(* CODESYS project jsontools.library
   DefaultNamespace: KOSTAL.AF2024.Core.JsonTools
   DocFormat: reStructuredText
   Description: Base functionalities to handle a json File
   Author: Frank Dümpelmann
   Title: KOSTAL.AF2024.Core.JsonTools
   Version: 1.0.0.0
   Company: KOSTAL GmbH & Co.KG
   Placeholder: KOSTAL.AF2024.Core.JsonTools

Project tree, tasks and I/O mapping:
  libraries: KOSTAL.AF2024.Core.Process, 1.0.0.0 (KOSTAL GmbH & Co.KG); KOSTAL.AF2024.Core.Settings, 1.0.0.0 (KOSTAL GmbH & Co.KG); KOSTAL.AF2024.Core.StringTools, 1.0.0.0 (KOSTAL GmbH & Co.KG); KOSTAL.AF2024.Core.System, 1.0.0.0 (KOSTAL GmbH & Co.KG); Tc2_Standard, 3.3.3.0 (Beckhoff Automation GmbH); Tc2_System, 3.6.2.0 (Beckhoff Automation GmbH); Tc2_Utilities, 3.5.2.0 (Beckhoff Automation GmbH); Tc3_IotBase, 3.3.2.0 (Beckhoff Automation GmbH); Tc3_JsonXml, 3.4.3.0 (Beckhoff Automation GmbH)
  0_Core/
    function block _FB_Core [ST]: _DocumentIsEmpty, _FBmain, _GetArrayElementByIndex, _GetArraySize, _GetDocument, _GetDocumentLenght, _NewDocument, FB_exit, FBmain
  1_Base/
    0_Protected/
      function block _FB_Base_PE [ST]: _ReadExtStorage, _ReadFileStorage, _FB_Main_EXT, _Step_ClearContent, _Step_CreateContent, _Step_Idle_EXT, _Step_ParseContent, _Step_ReadFile, _Step_ValidateFile, _Step_WriteFileAs, _Step_WriteFileVerification, _Step_Clear, _Step_failed, _Step_Finish, _Step_FinishFail, _Step_Idle, _Step_ValidateParameter, _WriteExtAsStorage, _wFV_a0_ChainFail, _wFV_a0_Finish, _wFV_a10_Origin, _wFV_a10_Read, _WriteFileAsStorage, _extStorageDefine, _FBmain, _PE_Ex_ReadExt, _PE_Ex_ReadFile, _PE_Ex_SaveFileAs, _PE_Ex_SaveToExtAs, _PE_Clear, _PE_FBmain
    1_Public/
      0_Fundamental/
        function block _FB_Base [ST]: Clear, FBmain, LinkExtStorage, extFileName, extFilePath, fullQualifiedFile, State, TimeOut
      1_DataSourceAccess/
        function block _FB_Base_RO [ST]: Ex_ReadExt, Ex_ReadFile
        function block _FB_Base_RW [ST]: Ex_SaveFileAs, Ex_SaveToExtAs, Retries
  DUT/
    data type E_THIS_CALLED
  PARSING/
    function block _FB_Parsing [ST]: PARSE_ARRAY, PARSE_BOOL, PARSE_BYTE, PARSE_DINT, PARSE_JSON, PARSE_LREAL, PARSE_MEMBER, PARSE_REAL, PARSE_STRING, PARSE_TIME, PARSE_UDINT, PARSE_ULINT
    function block _FB_Parsing_PE [ST]: _PARSE_ARRAY, _PARSE_BOOL, _PARSE_BYTE, _PARSE_DINT, _PARSE_JSON, _PARSE_LREAL, _PARSE_MEMBER, _PARSE_REAL, _PARSE_STRING, _PARSE_TIME, _PARSE_UDINT, _PARSE_ULINT
  Project Information/
    function F_GetCompany [ST]
    function F_GetTitle [ST]
    function F_GetVersion [ST]
  Storage/
    interface I_JsonStorage: Ex_Read, Ex_Write, LinkJsonParser, State
  Version/
    global variables Global_Version
*)

// DUT/E_THIS_CALLED
{attribute 'qualified_only'}
{attribute 'strict'}
TYPE E_THIS_CALLED :
(
	IDL := 0,
	FILE_READ,
	FILE_WRITE,
	WEB_READ,
	WEB_WRITE,
	CLEAR
);
END_TYPE

// Version/Global_Version
{attribute 'TcGenerated'}
{attribute 'no-analysis'}
{attribute 'linkalways'}
// This function has been automatically generated from the project information.
VAR_GLOBAL CONSTANT
	{attribute 'const_non_replaced'}
	stLibVersion_KOSTAL_AF2024_Core_JsonTools : ST_LibVersion := (iMajor := 1, iMinor := 0, iBuild := 0, iRevision := 0, nFlags := 0, sVersion := '1.0.0.0');
END_VAR

// 0_Core/_FB_Core
(*
	Use the FB_Core class if you want to use your own json data source.
	e.g. a STRING(4096) on a communication.
*)
FUNCTION_BLOCK ABSTRACT _FB_Core EXTENDS _FB_Parsing_PE

VAR
	
	_jDoc		: Tc3_IotBase.SJsonValue;	

	_concat	: Kostal_AF2024_Core_StringTools.FB_CONCAT;
	
END_VAR

VAR CONSTANT
	_EMPTY_DOC_LENGHT	: UDINT:= 5;
END_VAR

METHOD PROTECTED _DocumentIsEmpty : BOOL

_DocumentIsEmpty:= _parser.GetDocumentLength() <= _EMPTY_DOC_LENGHT;
END_METHOD

METHOD PROTECTED _FBmain : BOOL
;
END_METHOD

METHOD PROTECTED _GetArrayElementByIndex : Tc3_IotBase.SJsonValue
VAR_INPUT
	jContainer	: Tc3_IotBase.SJsonValue;
	Index				: UDINT;
	state				: REFERENCE TO KOSTAL_AF2024_Core_Settings.T_MaxString;		
END_VAR

VAR
	_state					: KOSTAL_AF2024_Core_Settings.T_MaxString;	
END_VAR
IF jContainer = 0 THEN _state:= "GetArraySize - jContainer Parameter is empty";	

ELSIF Index >= _parser.GetArraySize(jContainer) THEN	_state:= "GetArraySize - Index is out of range";

ELSE	_GetArrayElementByIndex:= _parser.GetArrayValueByIdx(jContainer, Index);

END_IF

IF __ISVALIDREF(state) THEN state:= _state;	END_IF
END_METHOD

METHOD PROTECTED _GetArraySize : UDINT;
VAR_INPUT
	jContainer	: Tc3_IotBase.SJsonValue;
	state				: REFERENCE TO KOSTAL_AF2024_Core_Settings.T_MaxString;		
END_VAR

VAR
	_state	: KOSTAL_AF2024_Core_Settings.T_MaxString;	
END_VAR
IF jContainer = 0 THEN _state:= "GetArraySize - jContainer Parameter is empty";	

ELSE	_GetArraySize:= _parser.GetArraySize(jContainer);
	
END_IF

IF __ISVALIDREF(state) THEN state:= _state;	END_IF
END_METHOD

(*
getDocument
===========

|return a Pointer >Tc3_IotBase.SJsonValue< to jason document
*)

METHOD PROTECTED _GetDocument : Tc3_IotBase.SJsonValue;
_GetDocument:= _jDoc;
END_METHOD

METHOD PROTECTED _GetDocumentLenght : UDINT;
VAR_INPUT
END_VAR
_GetDocumentLenght:= _parser.GetDocumentLength();
END_METHOD

(*
use in your _Step_CreateContent to start with an empty json File
*)
METHOD PROTECTED _NewDocument : BOOL

_parser.NewDocument();

_jDoc:= _parser.GetDocumentRoot();

_GetDocumentLenght();

_NewDocument:= _jDoc <> 0;
END_METHOD

METHOD FB_exit : BOOL
VAR_INPUT
	bInCopyCode : BOOL; // if TRUE, the exit method is called for exiting an instance that is copied afterwards (online change).
END_VAR

_NewDocument();
END_METHOD

METHOD PUBLIC FBmain
VAR_INPUT
END_VAR
;
END_METHOD

END_FUNCTION_BLOCK

// PARSING/_FB_Parsing_PE
(*
	Contains protected methods to parse various data types.
*)
FUNCTION_BLOCK ABSTRACT _FB_Parsing_PE

VAR
	_parser	: Tc3_JsonXml.FB_JsonDomParser;
END_VAR

(*
Returns the Json Array Element of jContainer
*)
METHOD PROTECTED _PARSE_ARRAY : Tc3_IotBase.SJsonValue;

VAR_INPUT
	jContainer	: Tc3_IotBase.SJsonValue;
	Member			: KOSTAL_AF2024_Core_Settings.T_MaxString_UTF8;	
	mustExist		: BOOL;
	state				: REFERENCE TO KOSTAL_AF2024_Core_Settings.T_MaxString_UTF8;		
END_VAR

VAR
	_J						:	Tc3_IotBase.SJsonValue;
	_state	: KOSTAL_AF2024_Core_Settings.T_MaxString_UTF8;	
END_VAR
_PARSE_ARRAY:= 0;
_state:= '';

IF jContainer = 0 																		THEN	_state:= Tc2_Standard.CONCAT(Member,  ';PARSE_ARRAY - jContainer Parameter is empty');	

ELSIF NOT _parser.HasMember(jContainer, Member)	THEN	_state:= Tc2_Standard.CONCAT(Member,  ';PARSE_ARRAY - no member');

ELSE

	_J:= _parser.FindMember(jContainer,	Member);

	IF _J = 0 										THEN 	_state:= Tc2_Standard.CONCAT(Member,  ';PARSE_ARRAY - no member');	
	ELSIF _parser.IsNull(_J)	THEN 	_state:= Tc2_Standard.CONCAT(Member,  ';PARSE_ARRAY - is NULL');	
	ELSE																_PARSE_ARRAY:= _J;
	END_IF

END_IF

IF __ISVALIDREF(state) THEN state:= _state;	END_IF
END_METHOD

(*
Returns a bool Value of jContainer
*)
METHOD PROTECTED _PARSE_BOOL : BOOL

VAR_INPUT
	jContainer	: Tc3_IotBase.SJsonValue;
	Member			: KOSTAL_AF2024_Core_Settings.T_MaxString_UTF8;	
	mustExist		: BOOL;
	state				: REFERENCE TO KOSTAL_AF2024_Core_Settings.T_MaxString_UTF8;		
END_VAR

VAR
	_J			:	Tc3_IotBase.SJsonValue;
	_state	: KOSTAL_AF2024_Core_Settings.T_MaxString_UTF8;	
END_VAR
_PARSE_BOOL:= FALSE; 
_state:= '';

IF jContainer = 0 THEN _state:= Tc2_Standard.CONCAT(Member,  ';PARSE_BOOL - jContainer Parameter is empty');

ELSIF NOT _parser.HasMember(jContainer, Member) THEN
	
	IF mustExist THEN	_state:= Tc2_Standard.CONCAT(Member,  ';PARSE_BOOL - no member');	END_IF

ELSE

	_J:= _parser.FindMember(jContainer,	Member);

	IF _J = 0 											THEN	IF mustExist	THEN	_state:= Tc2_Standard.CONCAT(Member,  ';PARSE_BOOL - no member');	END_IF
	ELSIF _parser.IsNull(_J)		THEN	IF mustExist	THEN	_state:= Tc2_Standard.CONCAT(Member,  ';PARSE_BOOL - is NULL');	END_IF
	ELSIF _parser.IsBool(_J)		THEN	_PARSE_BOOL:= _parser.GetBool(v:= _J);	
	ELSIF _parser.IsNumber(_J)	THEN	_PARSE_BOOL:=  UDINT_TO_BOOL(_parser.GetUint(_J));
	ELSIF _parser.IsString(_J)	THEN	_PARSE_BOOL:=  STRING_TO_BOOL(_parser.GetString(_J));
	ELSE																	IF mustExist 	THEN	_state:= Tc2_Standard.CONCAT(Member,  ';PARSE_BOOL - not BOOL');	END_IF
	END_IF

END_IF
	
IF __ISVALIDREF(state) THEN state:= _state;	END_IF
END_METHOD

(*
Returns a byte Value of jContainer
*)
METHOD PROTECTED _PARSE_BYTE : BYTE

VAR_INPUT
	jContainer	: Tc3_IotBase.SJsonValue;
	Member			: KOSTAL_AF2024_Core_Settings.T_MaxString_UTF8;	
	mustExist		: BOOL;
	state				: REFERENCE TO KOSTAL_AF2024_Core_Settings.T_MaxString_UTF8;		
END_VAR

VAR
	_J						:	Tc3_IotBase.SJsonValue;
	_state				: KOSTAL_AF2024_Core_Settings.T_MaxString_UTF8;	
END_VAR
_PARSE_BYTE:= 0; 
_state:= '';

IF jContainer = 0 THEN _state:= Tc2_Standard.CONCAT(Member,  ';PARSE_BYTE - jContainer Parameter is empty');

ELSIF NOT _parser.HasMember(jContainer, Member) THEN
	
	IF mustExist THEN	_state:= Tc2_Standard.CONCAT(Member,  ';PARSE_BYTE - no member');	END_IF

ELSE

	_J:= _parser.FindMember(jContainer,	Member);

	IF _J = 0 											THEN	IF mustExist	THEN	_state:= Tc2_Standard.CONCAT(Member,  ';PARSE_BYTE - no member');	END_IF
	ELSIF _parser.IsNull(_J)		THEN	IF mustExist	THEN	_state:= Tc2_Standard.CONCAT(Member,  ';PARSE_BYTE - is NULL');	END_IF
	ELSIF _parser.IsBool(_J)		THEN	_PARSE_BYTE:= 	BOOL_TO_BYTE(_parser.GetBool(v:= _J));	
	ELSIF _parser.IsNumber(_J)	THEN	_PARSE_BYTE:=  UDINT_TO_BYTE(_parser.GetUint(_J));
	ELSIF _parser.IsString(_J)	THEN	_PARSE_BYTE:=  STRING_TO_BYTE(_parser.GetString(_J));
	ELSE																	IF mustExist 	THEN	_state:= Tc2_Standard.CONCAT(Member,  ';PARSE_BYTE - not BYTE');	END_IF
	END_IF

END_IF
	
IF __ISVALIDREF(state) THEN state:= _state;	END_IF
END_METHOD

(*
Returns a DINT Value of jContainer
*)
METHOD PROTECTED _PARSE_DINT : DINT

VAR_INPUT
	jContainer	: Tc3_IotBase.SJsonValue;
	Member			: KOSTAL_AF2024_Core_Settings.T_MaxString_UTF8;	
	mustExist		: BOOL;
	state				: REFERENCE TO KOSTAL_AF2024_Core_Settings.T_MaxString_UTF8;		
END_VAR

VAR
	_J						:	Tc3_IotBase.SJsonValue;
	_state				: KOSTAL_AF2024_Core_Settings.T_MaxString_UTF8;	
END_VAR
_PARSE_DINT:= 0; 
_state:= '';

IF jContainer = 0 THEN _state:= Tc2_Standard.CONCAT(Member,  ';PARSE_DINT - jContainer Parameter is empty');

ELSIF NOT _parser.HasMember(jContainer, Member) THEN
	
	IF mustExist THEN	_state:= Tc2_Standard.CONCAT(Member,  ';PARSE_DINT - no member');	END_IF

ELSE

	_J:= _parser.FindMember(jContainer,	Member);

	IF _J = 0 											THEN	IF mustExist	THEN	_state:= Tc2_Standard.CONCAT(Member,  ';PARSE_DINT - no member');	END_IF
	ELSIF _parser.IsNull(_J)		THEN	IF mustExist	THEN	_state:= Tc2_Standard.CONCAT(Member,  ';PARSE_DINT - is NULL');	END_IF
	ELSIF _parser.IsBool(_J)		THEN	_PARSE_DINT:= 	BOOL_TO_DINT(_parser.GetBool(v:= _J));	
	ELSIF _parser.IsNumber(_J)	THEN	_PARSE_DINT:=  UDINT_TO_DINT(_parser.GetUint(_J));
	ELSIF _parser.IsString(_J)	THEN	_PARSE_DINT:=  STRING_TO_DINT(_parser.GetString(_J));
	ELSE																	IF mustExist 	THEN	_state:= Tc2_Standard.CONCAT(Member,  ';PARSE_DINT - not DINT');	END_IF
	END_IF

END_IF
	
IF __ISVALIDREF(state) THEN state:= _state;	END_IF
END_METHOD

(*
Returns the Json Element of jContainer
*)
METHOD PROTECTED _PARSE_JSON : Tc3_IotBase.SJsonValue;

VAR_INPUT
	jContainer	: Tc3_IotBase.SJsonValue;
	Member			: KOSTAL_AF2024_Core_Settings.T_MaxString_UTF8;	
	mustExist		: BOOL;
	state				: REFERENCE TO KOSTAL_AF2024_Core_Settings.T_MaxString_UTF8;		
END_VAR

VAR
	_J	:	Tc3_IotBase.SJsonValue;
	_state	: KOSTAL_AF2024_Core_Settings.T_MaxString_UTF8;	
END_VAR
_PARSE_JSON:= 0;
_state:= '';

IF jContainer = 0 																		THEN	_state:= Tc2_Standard.CONCAT(Member,  ';PARSE_JSON - jContainer Parameter is empty');	

ELSIF NOT _parser.HasMember(jContainer, Member)	THEN	_state:= Tc2_Standard.CONCAT(Member,  ';PARSE_JSON - no member');

ELSE

	_J:= _parser.FindMember(jContainer,	Member);

	IF _J = 0 									THEN 	_state:= Tc2_Standard.CONCAT(Member,  ';PARSE_JSON - no member');	
	ELSIF _parser.IsNull(_J)		THEN 	_state:= Tc2_Standard.CONCAT(Member,  ';PARSE_JSON - is NULL');	
	ELSE															_PARSE_JSON:= _J;
	END_IF

END_IF

IF __ISVALIDREF(state) THEN state:= _state;	END_IF
END_METHOD

(*
Returns a ULINT Value of jContainer
*)
METHOD PROTECTED _PARSE_LREAL : LREAL

VAR_INPUT
	jContainer	: Tc3_IotBase.SJsonValue;
	Member			: KOSTAL_AF2024_Core_Settings.T_MaxString_UTF8;	
	mustExist		: BOOL;
	state				: REFERENCE TO KOSTAL_AF2024_Core_Settings.T_MaxString_UTF8;		
END_VAR

VAR
	_J						:	Tc3_IotBase.SJsonValue;
	_state				: KOSTAL_AF2024_Core_Settings.T_MaxString_UTF8;	
END_VAR

_PARSE_LREAL:= LREAL#0; 

_state:= '';

IF jContainer = 0 THEN _state:= Tc2_Standard.CONCAT(Member,  ';PARSE_LREAL - jContainer Parameter is empty');

ELSIF NOT _parser.HasMember(jContainer, Member) THEN
	
	IF mustExist THEN	_state:= Tc2_Standard.CONCAT(Member,  ';PARSE_LREAL - no member');	END_IF

ELSE

	_J:= _parser.FindMember(jContainer,	Member);

	IF _J = 0 											THEN	IF mustExist	THEN	_state:= Tc2_Standard.CONCAT(Member,  ';PARSE_LREAL - no member');	END_IF
	ELSIF _parser.IsNull(_J)		THEN	IF mustExist	THEN	_state:= Tc2_Standard.CONCAT(Member,  ';PARSE_LREAL - is NULL');	END_IF
	ELSIF _parser.IsBool(_J)		THEN	_PARSE_LREAL:= 	BOOL_TO_LREAL(_parser.GetBool(v:= _J));	
	ELSIF _parser.IsNumber(_J)	THEN	_PARSE_LREAL:= 	_parser.GetDouble(_J);
	ELSIF _parser.IsString(_J)	THEN	_PARSE_LREAL:=	STRING_TO_LREAL(_parser.GetString(_J));
	ELSE																	IF mustExist 	THEN	_state:= Tc2_Standard.CONCAT(Member,  ';PARSE_LREAL - not BYTE');	END_IF
	END_IF

END_IF
	
IF __ISVALIDREF(state) THEN state:= _state;	END_IF
END_METHOD

(*
Returns the Json Element of jContainer
*)
METHOD PROTECTED _PARSE_MEMBER : Tc3_IotBase.SJsonValue;

VAR_INPUT
	jContainer	: Tc3_IotBase.SJsonValue;
	Member			: KOSTAL_AF2024_Core_Settings.T_MaxString_UTF8;	
	mustExist		: BOOL;
	state				: REFERENCE TO KOSTAL_AF2024_Core_Settings.T_MaxString_UTF8;		
END_VAR

VAR
	_J	:	Tc3_IotBase.SJsonValue;
	_state	: KOSTAL_AF2024_Core_Settings.T_MaxString_UTF8;	
END_VAR
_PARSE_MEMBER:= 0;
_state:= '';

IF jContainer = 0 																		THEN	_state:= Tc2_Standard.CONCAT(Member,  ';PARSE_JSON - jContainer Parameter is empty');	

ELSIF NOT _parser.HasMember(jContainer, Member)	THEN	_state:= Tc2_Standard.CONCAT(Member,  ';PARSE_JSON - no member');

ELSE

	_J:= _parser.FindMember(jContainer,	Member);

	IF _J = 0																	THEN 	_state:= Tc2_Standard.CONCAT(Member,  ';PARSE_JSON - no member');
	ELSIF		mustExist AND _parser.IsNull(_J)	THEN 	_state:= Tc2_Standard.CONCAT(Member,  ';PARSE_MEMBER - is NULL');	
	ELSE																						_PARSE_MEMBER:= _J;
	END_IF

END_IF

IF __ISVALIDREF(state) THEN state:= _state;	END_IF
END_METHOD

(*
Returns a ULINT Value of jContainer
*)
METHOD PROTECTED _PARSE_REAL : REAL

VAR_INPUT
	jContainer	: Tc3_IotBase.SJsonValue;
	Member			: KOSTAL_AF2024_Core_Settings.T_MaxString_UTF8;	
	mustExist		: BOOL;
	state				: REFERENCE TO KOSTAL_AF2024_Core_Settings.T_MaxString_UTF8;		
END_VAR

VAR
	_J						:	Tc3_IotBase.SJsonValue;
	_state				: KOSTAL_AF2024_Core_Settings.T_MaxString_UTF8;	
END_VAR

_PARSE_REAL:= REAL#0; 

_state:= '';

IF jContainer = 0 THEN _state:= Tc2_Standard.CONCAT(Member,  ';PARSE_REAL - jContainer Parameter is empty');

ELSIF NOT _parser.HasMember(jContainer, Member) THEN
	
	IF mustExist THEN	_state:= Tc2_Standard.CONCAT(Member,  ';PARSE_REAL - no member');	END_IF

ELSE

	_J:= _parser.FindMember(jContainer,	Member);

	IF _J = 0 											THEN	IF mustExist	THEN	_state:= Tc2_Standard.CONCAT(Member,  ';PARSE_REAL - no member');	END_IF
	ELSIF _parser.IsNull(_J)		THEN	IF mustExist	THEN	_state:= Tc2_Standard.CONCAT(Member,  ';PARSE_REAL - is NULL');	END_IF
	ELSIF _parser.IsBool(_J)		THEN	_PARSE_REAL:= 	BOOL_TO_REAL(_parser.GetBool(v:= _J));	
	ELSIF _parser.IsNumber(_J)	THEN	_PARSE_REAL:= 	LREAL_TO_REAL(_parser.GetDouble(_J));
	ELSIF _parser.IsString(_J)	THEN	_PARSE_REAL:=	STRING_TO_REAL(_parser.GetString(_J));
	ELSE																	IF mustExist 	THEN	_state:= Tc2_Standard.CONCAT(Member,  ';PARSE_REAL - not BYTE');	END_IF
	END_IF

END_IF
	
IF __ISVALIDREF(state) THEN state:= _state;	END_IF
END_METHOD

(*
Returns a STRING Value of jContainer
*)
METHOD PROTECTED _PARSE_STRING : KOSTAL_AF2024_Core_Settings.T_MaxString_UTF8

VAR_INPUT
	jContainer	: Tc3_IotBase.SJsonValue;
	Member			: KOSTAL_AF2024_Core_Settings.T_MaxString_UTF8;	
	mustExist		: BOOL;
	state				: REFERENCE TO KOSTAL_AF2024_Core_Settings.T_MaxString_UTF8;		
END_VAR

VAR
	_J						:	Tc3_IotBase.SJsonValue;
	_state				: KOSTAL_AF2024_Core_Settings.T_MaxString_UTF8;	
END_VAR
_PARSE_STRING:= ''; 
_state:= '';

IF jContainer = 0 THEN _state:= Tc2_Standard.CONCAT(Member,  ';PARSE_STRING - jContainer Parameter is empty');

ELSIF NOT _parser.HasMember(jContainer, Member) THEN
	
	IF mustExist THEN	_state:= Tc2_Standard.CONCAT(Member,  ';PARSE_STRING - no member');	END_IF

ELSE

	_J:= _parser.FindMember(jContainer,	Member);

	IF _J = 0 									THEN	IF mustExist		THEN	_state:= Tc2_Standard.CONCAT(Member,  ';PARSE_STRING - no member');	END_IF
	ELSIF _parser.IsNull(_J)		THEN	IF mustExist		THEN	_state:= Tc2_Standard.CONCAT(Member,  ';PARSE_STRING - is NULL');	END_IF
	ELSIF _parser.IsBool(_J)		THEN	_PARSE_STRING:= 	BOOL_TO_STRING(_parser.GetBool(v:= _J));	
	ELSIF _parser.IsNumber(_J)	THEN	_PARSE_STRING:=  UDINT_TO_STRING(_parser.GetUint(_J));
	ELSIF _parser.IsString(_J)	THEN	_PARSE_STRING:=  _parser.GetString(_J);
	ELSE				IF mustExist 		THEN	_state:= Tc2_Standard.CONCAT(Member,  ';PARSE_STRING - not STRING');	END_IF
	END_IF

END_IF
	
IF __ISVALIDREF(state) THEN state:= _state;	END_IF
END_METHOD

(*
Returns a TIME Value of jContainer
*)
METHOD PROTECTED _PARSE_TIME : TIME

VAR_INPUT
	jContainer	: Tc3_IotBase.SJsonValue;
	Member			: KOSTAL_AF2024_Core_Settings.T_MaxString_UTF8;	
	mustExist		: BOOL;
	state				: REFERENCE TO KOSTAL_AF2024_Core_Settings.T_MaxString_UTF8;		
END_VAR

VAR
	_J						:	Tc3_IotBase.SJsonValue;
	_num					: ULINT;
	_state				: KOSTAL_AF2024_Core_Settings.T_MaxString_UTF8;	
END_VAR
_PARSE_TIME:= T#0MS; 
_state:= '';

IF jContainer = 0 THEN _state:= Tc2_Standard.CONCAT(Member,  ';PARSE_TIME - jContainer Parameter is empty');

ELSIF NOT _parser.HasMember(jContainer, Member) THEN
	
	IF mustExist THEN	_state:= Tc2_Standard.CONCAT(Member,  ';PARSE_TIME - no member');	END_IF

ELSE

	_J:= _parser.FindMember(jContainer,	Member);

	IF _J = 0 									THEN	IF mustExist	THEN	_state:= Tc2_Standard.CONCAT(Member,  ';PARSE_TIME - no member');	END_IF
	ELSIF _parser.IsNull(_J)		THEN	IF mustExist	THEN	_state:= Tc2_Standard.CONCAT(Member,  ';PARSE_TIME - is NULL');	END_IF
	ELSIF _parser.IsNumber(_J)	THEN	_PARSE_TIME:=  ULINT_TO_TIME(_parser.GetUint(_J));
	ELSIF _parser.IsString(_J)	THEN	_PARSE_TIME:=  STRING_TO_TIME(_parser.GetString(_J));
	ELSE					IF mustExist 	THEN	_state:= Tc2_Standard.CONCAT(Member,  ';PARSE_TIME - not BYTE');	END_IF
	END_IF

END_IF
	
IF __ISVALIDREF(state) THEN state:= _state;	END_IF
END_METHOD

(*
Returns a UDINT Value of jContainer
*)
METHOD PROTECTED _PARSE_UDINT : UDINT

VAR_INPUT
	jContainer	: Tc3_IotBase.SJsonValue;
	Member			: KOSTAL_AF2024_Core_Settings.T_MaxString_UTF8;	
	mustExist		: BOOL;
	state				: REFERENCE TO KOSTAL_AF2024_Core_Settings.T_MaxString_UTF8;		
END_VAR

VAR
	_J						:	Tc3_IotBase.SJsonValue;
	_state				: KOSTAL_AF2024_Core_Settings.T_MaxString_UTF8;	
END_VAR
_PARSE_UDINT:= 0; 
_state:= '';

IF jContainer = 0 THEN _state:= Tc2_Standard.CONCAT(Member,  ';PARSE_UDINT - jContainer Parameter is empty');

ELSIF NOT _parser.HasMember(jContainer, Member) THEN
	
	IF mustExist THEN	_state:= Tc2_Standard.CONCAT(Member,  ';PARSE_UDINT - no member');	END_IF

ELSE

	_J:= _parser.FindMember(jContainer,	Member);

	IF _J = 0 									THEN	IF mustExist	THEN	_state:= Tc2_Standard.CONCAT(Member,  ';PARSE_UDINT - no member');	END_IF
	ELSIF _parser.IsNull(_J)		THEN	IF mustExist	THEN	_state:= Tc2_Standard.CONCAT(Member,  ';PARSE_UDINT - is NULL');	END_IF
	ELSIF _parser.IsBool(_J)		THEN	_PARSE_UDINT:= BOOL_TO_UDINT(_parser.GetBool(v:= _J));	
	ELSIF _parser.IsNumber(_J)	THEN	_PARSE_UDINT:= _parser.GetUint(_J);
	ELSIF _parser.IsString(_J)	THEN	_PARSE_UDINT:=  STRING_TO_UDINT(_parser.GetString(_J));
	ELSE					IF mustExist 	THEN	_state:= Tc2_Standard.CONCAT(Member,  ';PARSE_UDINT - not BYTE');	END_IF
	END_IF

END_IF
	
IF __ISVALIDREF(state) THEN state:= _state;	END_IF
END_METHOD

(*
Returns a ULINT Value of jContainer
*)
METHOD PROTECTED _PARSE_ULINT : ULINT

VAR_INPUT
	jContainer	: Tc3_IotBase.SJsonValue;
	Member			: KOSTAL_AF2024_Core_Settings.T_MaxString_UTF8;	
	mustExist		: BOOL;
	state				: REFERENCE TO KOSTAL_AF2024_Core_Settings.T_MaxString_UTF8;		
END_VAR

VAR
	_J						:	Tc3_IotBase.SJsonValue;
	_state				: KOSTAL_AF2024_Core_Settings.T_MaxString_UTF8;	
END_VAR
_PARSE_ULINT:= 0; 
_state:= '';

IF jContainer = 0 THEN _state:= Tc2_Standard.CONCAT(Member,  ';PARSE_ULINT - jContainer Parameter is empty');

ELSIF NOT _parser.HasMember(jContainer, Member) THEN
	
	IF mustExist THEN	_state:= Tc2_Standard.CONCAT(Member,  ';PARSE_ULINT - no member');	END_IF

ELSE

	_J:= _parser.FindMember(jContainer,	Member);

	IF _J = 0										THEN	IF mustExist	THEN	_state:= Tc2_Standard.CONCAT(Member,  ';PARSE_ULINT - no member');	END_IF
	ELSIF _parser.IsNull(_J)		THEN	IF mustExist	THEN	_state:= Tc2_Standard.CONCAT(Member,  ';PARSE_ULINT - is NULL');	END_IF
	ELSIF _parser.IsBool(_J)		THEN	_PARSE_ULINT:= BOOL_TO_ULINT(_parser.GetBool(v:= _J));	
	ELSIF _parser.IsNumber(_J)	THEN	_PARSE_ULINT:= _parser.GetUint64(_J);
	ELSIF _parser.IsString(_J)	THEN	_PARSE_ULINT:=  STRING_TO_ULINT(_parser.GetString(_J));
	ELSE					IF mustExist 	THEN	_state:= Tc2_Standard.CONCAT(Member,  ';PARSE_ULINT - not BYTE');	END_IF
	END_IF

END_IF
	
IF __ISVALIDREF(state) THEN state:= _state;	END_IF
END_METHOD

END_FUNCTION_BLOCK

// 1_Base/0_Protected/_FB_Base_PE
(*
	All needed methods and parameters are available as protected _..._PE templates
	make in inherating class available in puclic methods and parameters
*)
FUNCTION_BLOCK ABSTRACT _FB_Base_PE EXTENDS _FB_Core

VAR
	
	_Step				: KOSTAL_AF2024_Core_process.FB_processStep_Flow;

	_State	: KOSTAL_AF2024_Core_Process.T_plcState;

	_THIS_CALLED			: E_THIS_CALLED;
	_THIS_IN_PROCESS	: E_THIS_CALLED;

	_fullQualifiedFile	: KOSTAL_AF2024_Core_Settings.T_MaxString_UTF8;

	_ExecuteLoad	: BOOL;
	_LoadSuccess	: BOOL;

	_ExecuteSave	: BOOL;
	_SaveSuccess	: BOOL;

	
	_TimeOutTimer	: Tc2_Standard.TON;
	_TimeOut			: TIME:= T#5S;
	
	_iExtStorage	: I_JsonStorage;
	_extFileName	: KOSTAL_AF2024_Core_Settings.T_MaxString_UTF8;
	_extFilePath	: KOSTAL_AF2024_Core_Settings.T_MaxString_UTF8;
	
	{region 'write file verification'}
		_wFV_Step						: KOSTAL_AF2024_Core_process.FB_processStep_Flow;
		_wFV_Retries				: UINT:= 3;
		_wFV_RetriesCounter	: UINT;
		_wFV_FFE						: Tc2_Utilities.FB_EnumFindFileEntry;
		_wFV_ParserFileSize	: ULINT;
		_wFV_FileSize				: ULINT;
	{endregion}
	
	_ADDRESS_writeFailAs: INT;

END_VAR

VAR CONSTANT
	_ADDRESS_IDLE					: INT:= 0;
	_ADDRESS_SAVE_FILE_AS	: INT:= 100;
	_ADDRESS_CLEAR				: INT:= 200;
	_ADDRESS_FINISH_FAIL	: INT:= 300;
END_VAR

METHOD PROTECTED _ReadExtStorage
VAR_INPUT
END_VAR
IF _Step.toggle THEN	

	_TimeOutTimer(IN:= FALSE);	

	IF _iExtStorage = 0 THEN
		
		_State.clear();
		_State.finish:= TRUE;
		_State.fail:= TRUE;
		_State.description:= "web storage is not linked";
		
		_Step.set(_ADDRESS_FINISH_FAIL);

		RETURN;
	
	ELSIF NOT _iExtStorage.State.ready	THEN

		_State.clear();
		_State.finish:= TRUE;
		_State.fail:= TRUE;
		_State.description:= "web storage is not ready";
		
		_Step.set(_ADDRESS_FINISH_FAIL);

		RETURN;

	END_IF
	
END_IF


_TimeOutTimer(IN:= TRUE, PT:= _TimeOut);

IF _TimeOutTimer.Q THEN

	_State.clear();
	_State.finish:= TRUE;
	_State.fail:= TRUE;
	_State.description:= "File not able to read";

	_Step.set(_ADDRESS_FINISH_FAIL);

ELSIF NOT _iExtStorage.Ex_Read(_extFileName, _extFilePath) THEN	

	_State.clear();
	_State.busy:= TRUE;
	_State.description:= Tc2_Standard.WCONCAT("wait for web call accept;", _iExtStorage.State.description);

ELSIF NOT _iExtStorage.State.finish THEN	

	_State.clear();
	_State.busy:= TRUE;
	_State.description:= Tc2_Standard.WCONCAT("wait for web response;", _iExtStorage.State.description);

ELSIF NOT _iExtStorage.State.pass THEN	

	_State.clear();
	_State.finish:= TRUE;
	_State.fail:= TRUE;
	_State.description:= Tc2_Standard.WCONCAT("web call failed;", _iExtStorage.State.description);

	_Step.set(_ADDRESS_FINISH_FAIL);

ELSE	

	_jDoc:= _parser.GetDocumentRoot();
	_Step.INC();
			
END_IF
END_METHOD

METHOD PROTECTED _ReadFileStorage
VAR_INPUT
END_VAR


IF _Step.toggle THEN	_ExecuteLoad:= TRUE; _TimeOutTimer(IN:= FALSE);	END_IF

_TimeOutTimer(IN:= _ExecuteLoad, PT:= _TimeOut);

IF _ExecuteLoad THEN
	_LoadSuccess:= _parser.LoadDocumentFromFile(_fullQualifiedFile, _ExecuteLoad);
END_IF

IF _TimeOutTimer.Q THEN

	_State.clear();
	_State.finish:= TRUE;
	_State.fail:= TRUE;
	_State.description:= "File not able to read";

ELSIF _ExecuteLoad THEN	

	_State.description:= "Wait for LoadDocument Response";

ELSIF NOT _LoadSuccess THEN	

	_State.clear();
	_State.finish:= TRUE;
	_State.fail:= TRUE;
	_State.description:= "LoadDocument failed";
	
ELSE	

	_jDoc:= _parser.GetDocumentRoot();
	_Step.INC();
			
END_IF
END_METHOD

(*
	Overwrite to add your FBmain extension
*)
METHOD PROTECTED _FB_Main_EXT : BOOL
VAR_INPUT
END_VAR
END_METHOD

(*
	Overwrite to clear your data content before parse content
*)
METHOD PROTECTED _Step_ClearContent

_Step.INC();
END_METHOD

(*
	Overwrite to create your data content
*)
METHOD PROTECTED _Step_CreateContent

_Step.INC();
END_METHOD

(*
	Overwrite to add your Idle content here
*)
METHOD PROTECTED _Step_Idle_EXT : BOOL
VAR_INPUT
END_VAR

_Step_Idle_EXT:= FALSE;
END_METHOD

(*
	Overwrite to parse your data content
*)
METHOD PROTECTED _Step_ParseContent

_Step.INC();
END_METHOD

METHOD PROTECTED _Step_ReadFile
VAR_INPUT
END_VAR

IF 		_THIS_IN_PROCESS = E_THIS_CALLED.FILE_READ 	THEN	_ReadFileStorage();
ELSIF	_THIS_IN_PROCESS = E_THIS_CALLED.WEB_READ 	THEN	_ReadExtStorage();
ELSE

	_State.clear();
	_State.description:= Tc2_Standard.WCONCAT("no valid process in _Step_ReadFile; IN_PROCESS: ", INT_TO_WSTRING(_THIS_IN_PROCESS));
	_State.finish:= TRUE;
	_State.fail:= TRUE;
	_step.set(_ADDRESS_FINISH_FAIL);

END_IF
END_METHOD

METHOD PROTECTED _Step_ValidateFile
VAR_INPUT
END_VAR

_State.clear();
_State.finish:= TRUE;

IF _DocumentIsEmpty() THEN	

	_State.clear();
	_State.finish:= TRUE;
	_State.fail:= TRUE;
	_State.description:= "File not found or empty";

ELSE

	_Step.INC();

END_IF
END_METHOD

METHOD PROTECTED _Step_WriteFileAs
VAR_INPUT
END_VAR

_ADDRESS_writeFailAs:= _Step.actual;

IF 		_THIS_IN_PROCESS = E_THIS_CALLED.FILE_WRITE THEN	_WriteFileAsStorage();
ELSIF	_THIS_IN_PROCESS = E_THIS_CALLED.WEB_WRITE 	THEN	_WriteExtAsStorage();
ELSE

	_State.clear();
	_State.description:= Tc2_Standard.WCONCAT("no valid process in _Step_WriteFileAs; IN_PROCESS: ", INT_TO_WSTRING(_THIS_IN_PROCESS));
	_State.finish:= TRUE;
	_State.fail:= TRUE;
	_step.set(_ADDRESS_FINISH_FAIL);

END_IF
END_METHOD

METHOD PROTECTED _Step_WriteFileVerification

IF _THIS_IN_PROCESS <> E_THIS_CALLED.FILE_WRITE THEN	_Step.INC();
ELSE

	IF _Step.toggle	THEN	_wFV_Step.init();	END_IF
	
	_wFV_Step.Header();
	
	IF _wFV_Step.isActive(0)	THEN	_wFV_a10_Origin();	END_IF
	IF _wFV_Step.isActive(1)	THEN	_wFV_a10_Read();		END_IF
	IF _wFV_Step.isActive(2)	THEN	_wFV_a0_Finish();		END_IF
	
	IF _wFV_Step.NotFound()	THEN _wFV_a0_ChainFail();		END_IF

END_IF
END_METHOD

METHOD PROTECTED _Step_Clear
VAR_INPUT
END_VAR

_NewDocument();	

_Step.INC();
END_METHOD

METHOD PROTECTED _Step_failed
VAR_INPUT
END_VAR

_State.clear();
_State.finish:= TRUE;
_State.fail:= TRUE;

_concat.clear();
_concat.addContent("STEP Number ");
_concat.addContent(INT_TO_WSTRING(_Step.actual));
_concat.addContent(" does not exist - PLease call Support");

_State.description:= _concat.getResult();

_concat.clear();
END_METHOD

METHOD PROTECTED _Step_Finish : BOOL
VAR_INPUT
END_VAR

_State.clear();
_State.finish:= TRUE;
_State.pass:= TRUE;

_Step_Finish:= TRUE;
END_METHOD

METHOD PROTECTED _Step_FinishFail

VAR_INST
	_description	: KOSTAL_AF2024_Core_Settings.T_MaxString;
END_VAR

IF _Step.toggle THEN _description:= _State.description;	END_IF

_state.clear(); 
_state.finish := true;
_state.fail:= TRUE;

_state.description:= _description;
END_METHOD

METHOD PROTECTED _Step_Idle
VAR_INPUT
END_VAR

VAR
	_EmptyFile: KOSTAL_AF2024_Core_Settings.T_MaxString_UTF8;
END_VAR

IF _Step.toggle THEN
	
	_EmptyFile:= '';
	
	_ExecuteLoad:= FALSE;
	_LoadSuccess:= _parser.LoadDocumentFromFile(_EmptyFile, _ExecuteLoad);
	_LoadSuccess:= FALSE;

	_ExecuteSave:= FALSE;
	_SaveSuccess:= _parser.SaveDocumentToFile(_EmptyFile, _ExecuteSave);
	_SaveSuccess:= FALSE;
	
	_wFV_RetriesCounter:= UINT#0;

END_IF

IF _Step_Idle_EXT() THEN	; //Handle extended content

ELSIF _THIS_CALLED = E_THIS_CALLED.FILE_READ THEN

	_THIS_IN_PROCESS:= _THIS_CALLED;

	_NewDocument();
	_State.clear();
	_State.busy:= TRUE;
	_step.INC();


ELSIF _THIS_CALLED = E_THIS_CALLED.WEB_READ THEN

	_THIS_IN_PROCESS:= _THIS_CALLED;
	
	_NewDocument();
	_State.clear();
	_State.busy:= TRUE;
	_step.INC();



ELSIF _THIS_CALLED = E_THIS_CALLED.FILE_WRITE THEN

	_THIS_IN_PROCESS:= _THIS_CALLED;

	_State.clear();
	_State.busy:= TRUE;
	_step.set(_ADDRESS_SAVE_FILE_AS);


ELSIF _THIS_CALLED = E_THIS_CALLED.WEB_WRITE THEN

	_THIS_IN_PROCESS:= _THIS_CALLED;

	_State.clear();
	_State.busy:= TRUE;
	_step.set(_ADDRESS_SAVE_FILE_AS);



ELSIF _THIS_CALLED = E_THIS_CALLED.CLEAR THEN

	_THIS_IN_PROCESS:= _THIS_CALLED;

	_State.clear();
	_State.busy:= TRUE;
	_step.set(_ADDRESS_CLEAR);

ELSE

	_THIS_IN_PROCESS:= E_THIS_CALLED.IDL;	

	_State.clear();
	_State.ready:= TRUE;


END_IF
END_METHOD

METHOD PROTECTED _Step_ValidateParameter
VAR_INPUT
END_VAR

IF (_THIS_IN_PROCESS = E_THIS_CALLED.FILE_READ)
OR (_THIS_IN_PROCESS = E_THIS_CALLED.FILE_WRITE) 	
THEN

	IF _fullQualifiedFile = '' THEN	

		_State.clear();
		_State.finish:= TRUE;
		_State.fail:= TRUE;
		_State.description:= "fullQualifiedFile is empty";

	ELSE

		_Step.INC();
		
	END_IF

ELSIF (_THIS_IN_PROCESS = E_THIS_CALLED.WEB_READ)
OR 		(_THIS_IN_PROCESS = E_THIS_CALLED.WEB_WRITE) 	
THEN

	IF _extFileName = '' THEN	

		_State.clear();
		_State.finish:= TRUE;
		_State.fail:= TRUE;
		_State.description:= "webFileName is empty";

	ELSIF _extFilePath = '' THEN	

		_State.clear();
		_State.finish:= TRUE;
		_State.fail:= TRUE;
		_State.description:= "webFilePath is empty";

	ELSE

		_Step.INC();
		
	END_IF

ELSE
	
	_Step.INC();

END_IF
END_METHOD

METHOD PROTECTED _WriteExtAsStorage
VAR_INPUT
END_VAR
IF _Step.toggle THEN	

	_TimeOutTimer(IN:= FALSE);	

	IF _iExtStorage = 0 THEN
		
		_State.clear();
		_State.finish:= TRUE;
		_State.fail:= TRUE;
		_State.description:= "web storage is not linked";
		
		_Step.set(_ADDRESS_FINISH_FAIL);

		RETURN;
	
	ELSIF NOT _iExtStorage.State.ready	THEN

		_State.clear();
		_State.finish:= TRUE;
		_State.fail:= TRUE;
		_State.description:= "web storage is not ready";
		
		_Step.set(_ADDRESS_FINISH_FAIL);

		RETURN;

	END_IF
	
END_IF


_TimeOutTimer(IN:= TRUE, PT:= _TimeOut);

IF _TimeOutTimer.Q THEN

	_State.clear();
	_State.finish:= TRUE;
	_State.fail:= TRUE;
	_State.description:= "File not able to write";

	_Step.set(_ADDRESS_FINISH_FAIL);

ELSIF NOT _iExtStorage.Ex_Write(_extFileName, _extFilePath) THEN	

	_State.clear();
	_State.busy:= TRUE;
	_State.description:= Tc2_Standard.WCONCAT("wait for web call accept;", _iExtStorage.State.description);

ELSIF NOT _iExtStorage.State.finish THEN	

	_State.clear();
	_State.busy:= TRUE;
	_State.description:= Tc2_Standard.WCONCAT("wait for web response;", _iExtStorage.State.description);

ELSIF NOT _iExtStorage.State.pass THEN	

	_State.clear();
	_State.finish:= TRUE;
	_State.fail:= TRUE;
	_State.description:= Tc2_Standard.WCONCAT("web call failed;", _iExtStorage.State.description);

	_Step.set(_ADDRESS_FINISH_FAIL);

ELSE	

	_jDoc:= _parser.GetDocumentRoot();
	_Step.INC();
			
END_IF
END_METHOD

METHOD PROTECTED _wFV_a0_ChainFail
VAR
	_c: Kostal_AF2024_Core_StringTools.FB_CONCAT;
END_VAR

_c.clear();
_c.addContent("Step ");
_c.addContent(INT_TO_WSTRING(_wFV_Step.actual));
_c.addContent(" does not exist");

_State.clear();
_State.description:= _c.getResult();
_step.set(_ADDRESS_FINISH_FAIL);

_c.clear();
END_METHOD

METHOD PROTECTED _wFV_a0_Finish

_wFV_FFE(bExecute:= TRUE, eCmd:= Tc2_Utilities.E_EnumCmdType.eEnumCmd_Abort);
_wFV_FFE(bExecute:= FALSE);

_Step.INC();
END_METHOD

METHOD PROTECTED _wFV_a10_Origin

IF _Step.toggle	THEN	;	END_IF

_State.clear();
_State.busy:= TRUE;
_State.description:= "writeFile verification...";

_wFV_FFE(bExecute:= TRUE, eCmd:= Tc2_Utilities.E_EnumCmdType.eEnumCmd_Abort);
_wFV_FFE(bExecute:= FALSE);

_wFV_Step.INC();;
END_METHOD

METHOD PROTECTED _wFV_a10_Read

IF _wFV_Step.toggle THEN
	_wFV_FFE(bExecute:= TRUE, sPathName:= _fullQualifiedFile, sNetId:= '', eCmd:= Tc2_Utilities.E_EnumCmdType.eEnumCmd_First, tTimeout:= _TimeOut);
END_IF

_wFV_FFE(bExecute:= FALSE);

IF _Step.toggle	THEN	;	END_IF

_State.clear();

IF _wFV_FFE.bBusy	THEN

	_State.busy:= TRUE;
	_State.description:= "re-read written file";
	
ELSIF _wFV_FFE.bError	THEN

	IF _wFV_RetriesCounter >= _wFV_Retries	THEN
		
		_State.clear();
		_State.description:= "re-read written file - retries overflow";
		_step.set(_ADDRESS_FINISH_FAIL);
		
	ELSE
		
		_wFV_RetriesCounter:= _wFV_RetriesCounter + 1;

		_State.busy:= TRUE;
		_State.description:= "re-read written file failed - tryagain";
		_Step.set(_ADDRESS_writeFailAs);
		
	END_IF

ELSE
	
	_wFV_FileSize:= Tc2_Utilities.ULARGE_TO_ULINT(_wFV_FFE.stFindFile.fileSize);
	_wFV_ParserFileSize:= UDINT_TO_ULINT(_parser.GetDocumentLength());

	(*Parser size included the null-termination character - FileSize not*)
	IF (_wFV_FileSize + 1) <> _wFV_ParserFileSize	THEN	

		IF _wFV_RetriesCounter >= _wFV_Retries	THEN
			
			_State.clear();
			_State.description:= "re-read written file - size does not match - retries overflow";
			_step.set(_ADDRESS_FINISH_FAIL);
	
		ELSE
			
			_wFV_RetriesCounter:= _wFV_RetriesCounter + 1;
			_Step.set(_ADDRESS_writeFailAs);
			
		END_IF

	ELSE
	
		_wFV_RetriesCounter:= UINT#0;
		
		_wFV_Step.INC();;
	
	END_IF

END_IF
END_METHOD

METHOD PROTECTED _WriteFileAsStorage
VAR_INPUT
END_VAR


IF _Step.toggle THEN	_ExecuteSave:= TRUE;	_TimeOutTimer(IN:= FALSE);	END_IF

_TimeOutTimer(IN:= _ExecuteSave, PT:= _TimeOut);

IF _ExecuteSave THEN
	_SaveSuccess:= _parser.SaveDocumentToFile(_fullQualifiedFile, _ExecuteSave);
END_IF

IF _TimeOutTimer.Q THEN

	_State.clear();
	_State.finish:= TRUE;
	_State.fail:= TRUE;
	_State.description:= "File not able to write";

ELSIF _ExecuteSave THEN	

	_State.description:= "Wait for SaveDocument Response";

ELSIF NOT _SaveSuccess THEN	

	_State.clear();
	_State.finish:= TRUE;
	_State.fail:= TRUE;
	_State.description:= "SaveDocument failed";
			
ELSE	

	_step.INC();

END_IF
END_METHOD

METHOD PROTECTED _extStorageDefine
VAR_INPUT
END_VAR

IF _iExtStorage <> 0 THEN
	
	_iExtStorage.LinkJsonParser(_parser);
	
END_IF
END_METHOD

METHOD PROTECTED _FBmain : BOOL
_extStorageDefine();

IF _THIS_CALLED <> _THIS_IN_PROCESS AND _Step.actual <> 0 THEN	_Step.init();	END_IF
	
_Step.Header();

IF	_Step.isActive(_ADDRESS_IDLE)	THEN	_Step_Idle();	END_IF

//Read
IF	_Step.isActive(1)	THEN	_Step_ClearContent();				END_IF
IF	_Step.isActive(2)	THEN	_Step_ValidateParameter();	END_IF
IF	_Step.isActive(3)	THEN	_Step_ReadFile();						END_IF
IF	_Step.isActive(4)	THEN	_Step_ValidateFile();				END_IF
IF	_Step.isActive(5)	THEN	_Step_ParseContent();				END_IF
IF	_Step.isActive(6)	THEN	_Step_Finish();		END_IF

//Write
IF	_Step.isActive(_ADDRESS_SAVE_FILE_AS + 0)	THEN	_Step_ValidateParameter();			END_IF
IF	_Step.isActive(_ADDRESS_SAVE_FILE_AS + 1)	THEN	_Step_CreateContent();					END_IF
IF	_Step.isActive(_ADDRESS_SAVE_FILE_AS + 2)	THEN	_Step_WriteFileAs();						END_IF
IF	_Step.isActive(_ADDRESS_SAVE_FILE_AS + 3)	THEN	_Step_WriteFileVerification();	END_IF
IF	_Step.isActive(_ADDRESS_SAVE_FILE_AS + 4)	THEN	_Step_Finish();									END_IF

//Clear
IF	_Step.isActive(_ADDRESS_CLEAR)			THEN	_Step_Clear();				END_IF
IF	_Step.isActive(_ADDRESS_CLEAR + 1)	THEN	_Step_ClearContent();	END_IF
IF	_Step.isActive(_ADDRESS_CLEAR + 2)	THEN	_Step_Finish();				END_IF


//Finish - Failed
IF	_Step.isActive(_ADDRESS_FINISH_FAIL)	THEN	_Step_FinishFail();	END_IF



//Handle extended content
_FB_Main_EXT();


IF	_Step.NotFound() THEN	_Step_failed();	END_IF


_FBmain:= _THIS_CALLED = _THIS_IN_PROCESS;
END_METHOD

METHOD PROTECTED _PE_Ex_ReadExt : BOOL
VAR_INPUT
	FileName	: KOSTAL_AF2024_Core_Settings.T_MaxString_UTF8;	//Optional - if empty it will tried to use the stored Filename from Property WebFileName
	FilePath	: KOSTAL_AF2024_Core_Settings.T_MaxString_UTF8;	//Optional - if empty it will tried to use the stored Filename from Property WebFilePath
END_VAR
 
IF _THIS_CALLED = E_THIS_CALLED.IDL THEN

	_THIS_CALLED:= E_THIS_CALLED.WEB_READ;
	
	IF FileName <> '' THEN	_extFileName:= FileName;	END_IF
	IF FilePath <> '' THEN	_extFilePath:= FilePath;	END_IF

	_FBmain();
	
	_PE_Ex_ReadExt:= _THIS_CALLED = _THIS_IN_PROCESS;
	
ELSE
	
	_PE_Ex_ReadExt:= FALSE;
 
END_IF
END_METHOD

METHOD PROTECTED _PE_Ex_ReadFile : BOOL
VAR_INPUT
	full_Qualified_FileName	: KOSTAL_AF2024_Core_Settings.T_MaxString_UTF8;	//Optional - if empty it will tried to use the stored Filename from _fullQualifiedFileName
END_VAR
 
IF _THIS_CALLED = E_THIS_CALLED.IDL THEN

	_THIS_CALLED:= E_THIS_CALLED.FILE_READ;
	
	IF full_Qualified_FileName <> '' THEN	_fullQualifiedFile:= full_Qualified_FileName;	END_IF

	_FBmain();
	
	_PE_Ex_ReadFile:= _THIS_CALLED = _THIS_IN_PROCESS;

ELSE

	_PE_Ex_ReadFile:= FALSE;
 
END_IF
END_METHOD

METHOD PROTECTED _PE_Ex_SaveFileAs : BOOL
VAR_INPUT
	full_Qualified_FileName	: KOSTAL_AF2024_Core_Settings.T_MaxString_UTF8;	//Optional - if empty it will tried to use the stored Filename from _fullQualifiedFileName
END_VAR
 
IF _THIS_CALLED = E_THIS_CALLED.IDL THEN

	_THIS_CALLED:= E_THIS_CALLED.FILE_WRITE;
	
	IF full_Qualified_FileName <> '' THEN	_fullQualifiedFile:= full_Qualified_FileName;	END_IF

	_FBmain();

	_PE_Ex_SaveFileAs:= _THIS_CALLED = _THIS_IN_PROCESS;
	
ELSE
	
	_PE_Ex_SaveFileAs:= FALSE; 

END_IF
END_METHOD

METHOD PROTECTED _PE_Ex_SaveToExtAs : BOOL
VAR_INPUT
	FileName	: KOSTAL_AF2024_Core_Settings.T_MaxString_UTF8;	//Optional - if empty it will tried to use the stored Filename from Property WebFileName
	FilePath	: KOSTAL_AF2024_Core_Settings.T_MaxString_UTF8;	//Optional - if empty it will tried to use the stored Filename from Property WebFilePath
END_VAR
 
IF _THIS_CALLED = E_THIS_CALLED.IDL THEN

	_THIS_CALLED:= E_THIS_CALLED.WEB_WRITE;
	
	IF FileName <> ''	THEN	_extFileName:= FileName;	END_IF
	IF FilePath <> '' THEN	_extFilePath:= FilePath;	END_IF

	_FBmain();

	_PE_Ex_SaveToExtAs:= _THIS_CALLED = _THIS_IN_PROCESS;
	
ELSE

	_PE_Ex_SaveToExtAs:= FALSE;
	
END_IF
END_METHOD

METHOD PROTECTED _PE_Clear : BOOL

 
IF _THIS_CALLED = E_THIS_CALLED.IDL THEN

	_THIS_CALLED:= E_THIS_CALLED.CLEAR;

	_FBmain();

	_PE_Clear:= _THIS_CALLED = _THIS_IN_PROCESS;
 
END_IF
END_METHOD

METHOD PROTECTED _PE_FBmain


IF _THIS_CALLED = E_THIS_CALLED.IDL THEN
	_FBmain();
END_IF

_THIS_CALLED:= E_THIS_CALLED.IDL;
END_METHOD

END_FUNCTION_BLOCK

// Storage/I_JsonStorage
INTERFACE I_JsonStorage EXTENDS KOSTAL_AF2024_Core_System.I_Interface

METHOD Ex_Read : BOOL

VAR_INPUT
	FileName	: KOSTAL_AF2024_Core_Settings.T_MaxString_UTF8;
	FilePath	: KOSTAL_AF2024_Core_Settings.T_MaxString_UTF8;
END_VAR
END_METHOD

METHOD Ex_Write : BOOL

VAR_INPUT
	FileName	: KOSTAL_AF2024_Core_Settings.T_MaxString_UTF8;
	FilePath	: KOSTAL_AF2024_Core_Settings.T_MaxString_UTF8;
END_VAR
END_METHOD

METHOD PUBLIC LinkJsonParser
VAR_INPUT
	rJsonParser	: REFERENCE TO Tc3_JsonXml.FB_JsonDomParserBase;
END_VAR
END_METHOD

PROPERTY State : KOSTAL_AF2024_Core_Process.I_T_plcState
GET
END_GET
END_PROPERTY

END_INTERFACE

// 1_Base/1_Public/0_Fundamental/_FB_Base
(*
	FB_RootBase PUBLIC
	Fundamental methods and parameters are as public available.
	Add further required methods and properties to your inheriting class.
*)
FUNCTION_BLOCK ABSTRACT _FB_Base EXTENDS _FB_Base_PE

METHOD PUBLIC Clear : BOOL

SUPER^._PE_Clear();
END_METHOD

METHOD PUBLIC FBmain
 
SUPER^._PE_FBmain();
END_METHOD

METHOD PUBLIC LinkExtStorage
VAR_INPUT
	IN	: I_JsonStorage;
END_VAR

_iExtStorage	:= IN;
END_METHOD

PROPERTY PUBLIC extFileName : KOSTAL_AF2024_Core_Settings.T_MaxString_UTF8
GET

extFileName:= _extFileName;
END_GET
SET

_extFileName:= extFileName;
END_SET
END_PROPERTY

PROPERTY PUBLIC extFilePath : KOSTAL_AF2024_Core_Settings.T_MaxString_UTF8
GET

extFilePath:= _extFilePath;
END_GET
SET

_extFilePath:= extFilePath;
END_SET
END_PROPERTY

PROPERTY PUBLIC fullQualifiedFile : KOSTAL_AF2024_Core_Settings.T_MaxString_UTF8
GET

fullQualifiedFile:= _fullQualifiedFile;
END_GET
SET

_fullQualifiedFile:= fullQualifiedFile;
END_SET
END_PROPERTY

PROPERTY PUBLIC State : KOSTAL_AF2024_Core_Process.I_T_plcState
GET

State:= _State;
END_GET
END_PROPERTY

PROPERTY PUBLIC TimeOut : TIME
GET

TimeOut:= _TimeOut;
END_GET
SET

_TimeOut:= TimeOut;
END_SET
END_PROPERTY

END_FUNCTION_BLOCK

// 1_Base/1_Public/1_DataSourceAccess/_FB_Base_RO
(*
	FB_RootBase PUBLIC
	In addition to the functions of the FB_Base class, 
	the public methods for reading a source from a file 
	and an external data source are provided here.
*)
FUNCTION_BLOCK ABSTRACT _FB_Base_RO EXTENDS _FB_Base

METHOD PUBLIC Ex_ReadExt : BOOL
VAR_INPUT
	FileName	: KOSTAL_AF2024_Core_Settings.T_MaxString_UTF8;	//Optional - if empty it will tried to use the stored Filename from Property WebFileName
	FilePath	: KOSTAL_AF2024_Core_Settings.T_MaxString_UTF8;	//Optional - if empty it will tried to use the stored Filename from Property WebFilePath
END_VAR
Ex_ReadExt:= _PE_Ex_ReadExt(FileName, FilePath);
END_METHOD

METHOD PUBLIC Ex_ReadFile : BOOL
VAR_INPUT
	full_Qualified_FileName	: KOSTAL_AF2024_Core_Settings.T_MaxString_UTF8;	//Optional - if empty it will tried to use the stored Filename from _fullQualifiedFileName
END_VAR
Ex_ReadFile:= _PE_Ex_ReadFile(full_Qualified_FileName);
END_METHOD

END_FUNCTION_BLOCK

// 1_Base/1_Public/1_DataSourceAccess/_FB_Base_RW
(*
	In addition to the functions of the FB_Base_RO class, 
	the public methods for writing to a file 
	and to an external data source are provided here.
*)
FUNCTION_BLOCK ABSTRACT _FB_Base_RW EXTENDS _FB_Base_RO

METHOD PUBLIC Ex_SaveFileAs : BOOL
VAR_INPUT
	full_Qualified_FileName	: KOSTAL_AF2024_Core_Settings.T_MaxString_UTF8;	//Optional - if empty it will tried to use the stored Filename from _fullQualifiedFileName
END_VAR
Ex_SaveFileAs:= _PE_Ex_SaveFileAs(full_Qualified_FileName);
END_METHOD

METHOD PUBLIC Ex_SaveToExtAs : BOOL
VAR_INPUT
	FileName	: KOSTAL_AF2024_Core_Settings.T_MaxString_UTF8;	//Optional - if empty it will tried to use the stored Filename from Property WebFileName
	FilePath	: KOSTAL_AF2024_Core_Settings.T_MaxString_UTF8;	//Optional - if empty it will tried to use the stored Filename from Property WebFilePath
END_VAR
Ex_SaveToExtAs:= _PE_Ex_SaveToExtAs(FileName, FilePath);
END_METHOD

(*Contains the number of retries allowed for write attempts. *)
PROPERTY PUBLIC Retries : UINT
GET

Retries:= _wFV_Retries;
END_GET
SET

_wFV_Retries:= Retries;
END_SET
END_PROPERTY

END_FUNCTION_BLOCK

// PARSING/_FB_Parsing
(*
	Contains the public methods of the protected methods of the FB_Parsing_Root base class.
*)
FUNCTION_BLOCK PUBLIC _FB_Parsing EXTENDS _FB_Parsing_PE

(*
Returns the Json Array Element of jContainer
*)
METHOD PUBLIC PARSE_ARRAY : Tc3_IotBase.SJsonValue;

VAR_INPUT
	jContainer	: Tc3_IotBase.SJsonValue;
	Member			: KOSTAL_AF2024_Core_Settings.T_MaxString_UTF8;	
	mustExist		: BOOL;
	state				: REFERENCE TO KOSTAL_AF2024_Core_Settings.T_MaxString_UTF8;		
END_VAR

PARSE_ARRAY:= _PARSE_ARRAY(jContainer, Member, mustExist, state);
END_METHOD

(*
Returns a bool Value of jContainer
*)
METHOD PUBLIC PARSE_BOOL : BOOL

VAR_INPUT
	jContainer	: Tc3_IotBase.SJsonValue;
	Member			: KOSTAL_AF2024_Core_Settings.T_MaxString_UTF8;	
	mustExist		: BOOL;
	state				: REFERENCE TO KOSTAL_AF2024_Core_Settings.T_MaxString_UTF8;		
END_VAR

PARSE_BOOL:= _PARSE_BOOL(jContainer, Member, mustExist, state);
END_METHOD

(*
Returns a byte Value of jContainer
*)
METHOD PUBLIC PARSE_BYTE : BYTE

VAR_INPUT
	jContainer	: Tc3_IotBase.SJsonValue;
	Member			: KOSTAL_AF2024_Core_Settings.T_MaxString_UTF8;	
	mustExist		: BOOL;
	state				: REFERENCE TO KOSTAL_AF2024_Core_Settings.T_MaxString_UTF8;		
END_VAR

PARSE_BYTE:= _PARSE_BYTE(jContainer, Member, mustExist, state);
END_METHOD

(*
Returns a DINT Value of jContainer
*)
METHOD PUBLIC PARSE_DINT : DINT

VAR_INPUT
	jContainer	: Tc3_IotBase.SJsonValue;
	Member			: KOSTAL_AF2024_Core_Settings.T_MaxString_UTF8;	
	mustExist		: BOOL;
	state				: REFERENCE TO KOSTAL_AF2024_Core_Settings.T_MaxString_UTF8;		
END_VAR

PARSE_DINT:= _PARSE_DINT(jContainer, Member, mustExist, state);
END_METHOD

(*
Returns the Json Element of jContainer
*)
METHOD PUBLIC PARSE_JSON : Tc3_IotBase.SJsonValue;

VAR_INPUT
	jContainer	: Tc3_IotBase.SJsonValue;
	Member			: KOSTAL_AF2024_Core_Settings.T_MaxString_UTF8;	
	mustExist		: BOOL;
	state				: REFERENCE TO KOSTAL_AF2024_Core_Settings.T_MaxString_UTF8;		
END_VAR


PARSE_JSON:= _PARSE_JSON(jContainer, Member, mustExist, state);
END_METHOD

(*
Returns a ULINT Value of jContainer
*)
METHOD PUBLIC PARSE_LREAL : LREAL

VAR_INPUT
	jContainer	: Tc3_IotBase.SJsonValue;
	Member			: KOSTAL_AF2024_Core_Settings.T_MaxString_UTF8;	
	mustExist		: BOOL;
	state				: REFERENCE TO KOSTAL_AF2024_Core_Settings.T_MaxString_UTF8;		
END_VAR

PARSE_LREAL:= _PARSE_LREAL(jContainer, Member, mustExist, state);
END_METHOD

(*
Returns the Json Element of jContainer
*)
METHOD PUBLIC PARSE_MEMBER : Tc3_IotBase.SJsonValue;

VAR_INPUT
	jContainer	: Tc3_IotBase.SJsonValue;
	Member			: KOSTAL_AF2024_Core_Settings.T_MaxString_UTF8;	
	mustExist		: BOOL;
	state				: REFERENCE TO KOSTAL_AF2024_Core_Settings.T_MaxString_UTF8;		
END_VAR


PARSE_MEMBER:= _PARSE_MEMBER(jContainer, Member, mustExist, state);
END_METHOD

(*
Returns a ULINT Value of jContainer
*)
METHOD PUBLIC PARSE_REAL : REAL

VAR_INPUT
	jContainer	: Tc3_IotBase.SJsonValue;
	Member			: KOSTAL_AF2024_Core_Settings.T_MaxString_UTF8;	
	mustExist		: BOOL;
	state				: REFERENCE TO KOSTAL_AF2024_Core_Settings.T_MaxString_UTF8;		
END_VAR

PARSE_REAL:= _PARSE_REAL(jContainer, Member, mustExist, state);
END_METHOD

(*
Returns a STRING Value of jContainer
*)
METHOD PUBLIC PARSE_STRING : KOSTAL_AF2024_Core_Settings.T_MaxString_UTF8

VAR_INPUT
	jContainer	: Tc3_IotBase.SJsonValue;
	Member			: KOSTAL_AF2024_Core_Settings.T_MaxString_UTF8;	
	mustExist		: BOOL;
	state				: REFERENCE TO KOSTAL_AF2024_Core_Settings.T_MaxString_UTF8;		
END_VAR

PARSE_STRING:= _PARSE_STRING(jContainer, Member, mustExist, state);
END_METHOD

(*
Returns a TIME Value of jContainer
*)
METHOD PUBLIC PARSE_TIME : TIME

VAR_INPUT
	jContainer	: Tc3_IotBase.SJsonValue;
	Member			: KOSTAL_AF2024_Core_Settings.T_MaxString_UTF8;	
	mustExist		: BOOL;
	state				: REFERENCE TO KOSTAL_AF2024_Core_Settings.T_MaxString_UTF8;		
END_VAR


PARSE_TIME:= _PARSE_TIME(jContainer, Member, mustExist, state);
END_METHOD

(*
Returns a UDINT Value of jContainer
*)
METHOD PUBLIC PARSE_UDINT : UDINT

VAR_INPUT
	jContainer	: Tc3_IotBase.SJsonValue;
	Member			: KOSTAL_AF2024_Core_Settings.T_MaxString_UTF8;	
	mustExist		: BOOL;
	state				: REFERENCE TO KOSTAL_AF2024_Core_Settings.T_MaxString_UTF8;		
END_VAR

PARSE_UDINT:= _PARSE_UDINT(jContainer, Member, mustExist, state);
END_METHOD

(*
Returns a ULINT Value of jContainer
*)
METHOD PUBLIC PARSE_ULINT : ULINT

VAR_INPUT
	jContainer	: Tc3_IotBase.SJsonValue;
	Member			: KOSTAL_AF2024_Core_Settings.T_MaxString_UTF8;	
	mustExist		: BOOL;
	state				: REFERENCE TO KOSTAL_AF2024_Core_Settings.T_MaxString_UTF8;		
END_VAR

PARSE_ULINT:= _PARSE_ULINT(jContainer, Member, mustExist, state);
END_METHOD

END_FUNCTION_BLOCK

// Project Information/F_GetCompany
// This function has been automatically generated from the project information.
{attribute 'signature_flag' := '1073741824'}
{attribute 'TcGenerated'}
{attribute 'no-analysis'}
FUNCTION F_GetCompany : WSTRING
VAR_INPUT
	
END_VAR

F_GetCompany := "KOSTAL GmbH & Co.KG";

END_FUNCTION

// Project Information/F_GetTitle
// This function has been automatically generated from the project information.
{attribute 'signature_flag' := '1073741824'}
{attribute 'TcGenerated'}
{attribute 'no-analysis'}
FUNCTION F_GetTitle : WSTRING
VAR_INPUT
	
END_VAR

F_GetTitle := "KOSTAL.AF2024.Core.JsonTools";

END_FUNCTION

// Project Information/F_GetVersion
// This function has been automatically generated from the project information.
{attribute 'signature_flag' := '1073741824'}
{attribute 'TcGenerated'}
{attribute 'no-analysis'}
FUNCTION F_GetVersion : ST_LibVersion
VAR_INPUT
	
END_VAR

F_GetVersion.iMajor := 1;
F_GetVersion.iMinor := 0;
F_GetVersion.iBuild := 0;
F_GetVersion.iRevision := 0;
F_GetVersion.sVersion := '1.0.0.0';
F_GetVersion.nFlags := 0;

END_FUNCTION
